FUNCTION_BLOCK PalletAvailable (* Composite Function Block Type *)
  (* Standard: 61499-2 *)
  (* Version 0.0, 7/2/2026, template *)
  PACKAGE Main;
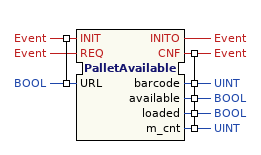
  EVENT_INPUT
    INIT WITH URL; (* Initialization Request *)
    REQ; (* Normal Execution Request *)
  END_EVENT
  EVENT_OUTPUT
    INITO; (* Initialization Confirm *)
    CNF WITH barcode, available, loaded, m_cnt; (* Execution Confirmation *)
  END_EVENT
  VAR_INPUT
    URL : BOOL; (* Input event qualifier *)
  END_VAR
  VAR_OUTPUT
    barcode : UINT; (* Output event qualifier *)
    available : BOOL;
    loaded : BOOL;
    m_cnt : UINT;
  END_VAR
END_FUNCTION_BLOCK
